(* IEC 61131-3 sources: PLCGen/codesys_service/bank/st_part4, 20 files *)

(* ---- E01_Filling.st ---- *)
(* Q01 Automated Filling Line Control - reference solution for test-case validation *)
FUNCTION_BLOCK E01_Filling
VAR_INPUT
    bottleSensor          : BOOL;
    cleaningConfirmButton : BOOL;
    fillingConfirmButton  : BOOL;
    cappingConfirmButton  : BOOL;
    packingConfirmButton  : BOOL;
    finishedButton        : BOOL;
END_VAR
VAR_OUTPUT
    Pump_Motor       : BOOL;
    Filling_Valve    : BOOL;
    Capping_Machine  : BOOL;
    Packing_Machine  : BOOL;
    Completion_Light : BOOL;
END_VAR
VAR
    step : INT := 0;   (* 0 idle, 1 cleaning, 2 filling, 3 capping, 4 packing, 5 done *)
    prevBottle      : BOOL;
    prevCleaning    : BOOL;
    prevFilling     : BOOL;
    prevCapping     : BOOL;
    prevPacking     : BOOL;
    prevFinished    : BOOL;
END_VAR

(* confirmation is edge-triggered: a button that is already held when its
   step is reached has no rising edge and must not confirm the step *)
IF step = 0 AND bottleSensor AND NOT prevBottle THEN
    step := 1;
ELSIF step = 1 AND cleaningConfirmButton AND NOT prevCleaning THEN
    step := 2;
ELSIF step = 2 AND fillingConfirmButton AND NOT prevFilling THEN
    step := 3;
ELSIF step = 3 AND cappingConfirmButton AND NOT prevCapping THEN
    step := 4;
ELSIF step = 4 AND packingConfirmButton AND NOT prevPacking THEN
    step := 5;
ELSIF step = 5 AND finishedButton AND NOT prevFinished THEN
    step := 0;
END_IF;

Pump_Motor       := step = 1;
Filling_Valve    := step = 2;
Capping_Machine  := step = 3;
Packing_Machine  := step = 4;
Completion_Light := step = 5;

prevBottle   := bottleSensor;
prevCleaning := cleaningConfirmButton;
prevFilling  := fillingConfirmButton;
prevCapping  := cappingConfirmButton;
prevPacking  := packingConfirmButton;
prevFinished := finishedButton;

(* ---- E02_DualEdge.st ---- *)
(* Q02 Dual-Word Edge Detection - reference solution *)
FUNCTION_BLOCK E02_DualEdge
VAR_INPUT
    value : DWORD;
END_VAR
VAR_OUTPUT
    hasChanged      : BOOL;
    hasRisingEdges  : BOOL;
    risingBits      : DWORD;
    noOfRisingBits  : USINT;
    hasFallingEdges : BOOL;
    fallingBits     : DWORD;
    noOfFallingBits : USINT;
END_VAR
VAR
    prev : DWORD;
    i    : INT;
    r    : DWORD;
    f    : DWORD;
END_VAR

risingBits  := value AND NOT prev;
fallingBits := prev AND NOT value;
hasChanged  := value <> prev;
hasRisingEdges  := risingBits <> 0;
hasFallingEdges := fallingBits <> 0;

(* popcount without SHL: shift right by division, which keeps the
   implementation portable and works in the simulator *)
r := risingBits;
f := fallingBits;
noOfRisingBits  := 0;
noOfFallingBits := 0;
FOR i := 0 TO 31 DO
    IF (r MOD 2) <> 0 THEN
        noOfRisingBits := noOfRisingBits + 1;
    END_IF;
    IF (f MOD 2) <> 0 THEN
        noOfFallingBits := noOfFallingBits + 1;
    END_IF;
    r := r / 2;
    f := f / 2;
END_FOR;

prev := value;

(* ---- E03_Hysteresis.st ---- *)
(* Q03 Alarm Handling - reference solution (used only to validate the test cases)
   Note: status codes are written in decimal (32769 = 16#8001, 32770 = 16#8002)
   because the offline simulator (st_sim) does not support typed literals. *)
FUNCTION_BLOCK E03_Hysteresis
VAR_INPUT
    Value      : REAL;
    hiLevel    : REAL;
    loLevel    : REAL;
    hystWindow : REAL;
END_VAR
VAR_OUTPUT
    hiAlarm : BOOL;
    loAlarm : BOOL;
    error   : BOOL;
    status  : WORD;
END_VAR

IF loLevel >= hiLevel THEN
    error  := TRUE;
    status := 32769;
ELSIF hystWindow >= hiLevel - loLevel THEN
    error  := TRUE;
    status := 32770;
ELSE
    error  := FALSE;
    status := 0;
    (* high alarm with hysteresis *)
    IF Value > hiLevel THEN
        hiAlarm := TRUE;
    ELSIF Value < hiLevel - hystWindow THEN
        hiAlarm := FALSE;
    END_IF;
    (* low alarm with hysteresis *)
    IF Value < loLevel THEN
        loAlarm := TRUE;
    ELSIF Value > loLevel + hystWindow THEN
        loAlarm := FALSE;
    END_IF;
END_IF;

(* ---- E04_JamPump.st ---- *)
(* Q04 Jam Pump Debouncing and Runtime Maintenance - reference solution
   Unit convention: TIME inputs in ms, LTIME output in ns (IEC 61131-3). *)
FUNCTION_BLOCK E04_JamPump
VAR_INPUT
    VISCOSITY_OK    : BOOL;
    PASTE_E_STOP_NC : BOOL;
    DebounceTime    : TIME;
    CycleTime       : TIME;
END_VAR
VAR_OUTPUT
    VFD_RUN          : BOOL;
    PUMP_MAINT_DUE   : BOOL;
    PUMP_RUNTIME_ACC : LTIME;
END_VAR
VAR
    debT    : TON;     (* real elapsed time, scan-clock driven *)
    accMs   : ULINT;   (* ms, per the team convention *)
END_VAR

(* VISCOSITY_OK must hold continuously for DebounceTime (real elapsed time) *)
debT(IN := VISCOSITY_OK AND PASTE_E_STOP_NC, PT := DebounceTime);
VFD_RUN := debT.Q AND PASTE_E_STOP_NC;

IF VFD_RUN THEN
    accMs := accMs + UDINT_TO_ULINT(TIME_TO_UDINT(CycleTime));
    PUMP_RUNTIME_ACC := ULINT_TO_LTIME(accMs);
END_IF;

IF accMs >= 1800000000 THEN   (* 500 h in ms *)
    PUMP_MAINT_DUE := TRUE;
END_IF;

(* ---- E05_WeldGap.st ---- *)
(* Q05 Weld Gap Alarm and Startup Inhibition - reference solution *)
FUNCTION_BLOCK E05_WeldGap
VAR_INPUT
    Gap_Exceeded   : BOOL;
    Weld_E_Stop_NC : BOOL;
    DebounceTime   : TIME;
END_VAR
VAR_OUTPUT
    Operator_Alert        : BOOL;
    Weld_Soft_Start_Active: BOOL;
END_VAR
VAR
    initTimer : TON;
    debTimer  : TON;
    initDone  : BOOL;
END_VAR

initTimer(IN := Weld_E_Stop_NC AND NOT initDone, PT := T#5S);
IF initTimer.Q THEN
    initDone := TRUE;
END_IF;

IF NOT Weld_E_Stop_NC THEN
    Operator_Alert := FALSE;
    Weld_Soft_Start_Active := FALSE;
    debTimer(IN := FALSE, PT := DebounceTime);
ELSIF NOT initDone THEN
    Operator_Alert := FALSE;
    Weld_Soft_Start_Active := TRUE;
    debTimer(IN := FALSE, PT := DebounceTime);
ELSE
    Weld_Soft_Start_Active := FALSE;
    debTimer(IN := Gap_Exceeded, PT := DebounceTime);
    Operator_Alert := debTimer.Q;
END_IF;

(* ---- E06_Blower.st ---- *)
(* Q06 Aeration Blower Delayed Start - reference solution *)
FUNCTION_BLOCK E06_Blower
VAR_INPUT
    DO_LOW               : BOOL;
    AERATION_E_STOP_NC   : BOOL;
END_VAR
VAR_OUTPUT
    BLOWER_RUN                  : BOOL;
    AERATION_BLOWER_CYCLE_COUNT : UINT;
END_VAR
VAR
    startTimer : TON;
    prevRun    : BOOL;
END_VAR

startTimer(IN := DO_LOW AND AERATION_E_STOP_NC, PT := T#5S);
BLOWER_RUN := startTimer.Q;

IF BLOWER_RUN AND NOT prevRun THEN
    AERATION_BLOWER_CYCLE_COUNT := AERATION_BLOWER_CYCLE_COUNT + 1;
END_IF;
prevRun := BLOWER_RUN;

(* ---- H01_Proportion.st ---- *)
(* Q15 Material Proportioning Process Control - reference solution for test-case validation *)
FUNCTION_BLOCK H01_Proportion
VAR_INPUT
    estop           : BOOL;
    opeMode         : BOOL;
    valveAStart     : BOOL;
    valveBStart     : BOOL;
    valveCStart     : BOOL;
    valveDStart     : BOOL;
    mixMotorStart   : BOOL;
    autoStart       : BOOL;
    processMode     : BOOL;
    levelSensor     : INT;
    mixMotorComplete: BOOL;
END_VAR
VAR_OUTPUT
    valveARun   : BOOL;
    valveBRun   : BOOL;
    valveCRun   : BOOL;
    valveDRun   : BOOL;
    mixMotorRun : BOOL;
END_VAR
VAR
    step : INT := 0;
    pA : BOOL;
    pB : BOOL;
    pC : BOOL;
    pD : BOOL;
    pM : BOOL;
END_VAR

IF NOT estop THEN
    valveARun := FALSE;
    valveBRun := FALSE;
    valveCRun := FALSE;
    valveDRun := FALSE;
    mixMotorRun := FALSE;
    step := 0;
ELSIF NOT opeMode THEN
    step := 0;
    IF valveAStart AND NOT pA THEN valveARun := NOT valveARun; END_IF;
    IF valveBStart AND NOT pB THEN valveBRun := NOT valveBRun; END_IF;
    IF valveCStart AND NOT pC THEN valveCRun := NOT valveCRun; END_IF;
    IF valveDStart AND NOT pD THEN valveDRun := NOT valveDRun; END_IF;
    IF mixMotorStart AND NOT pM THEN mixMotorRun := NOT mixMotorRun; END_IF;
ELSE
    IF step = 0 THEN
        valveARun := FALSE;
    valveBRun := FALSE;
    valveCRun := FALSE;
    valveDRun := FALSE;
    mixMotorRun := FALSE;
        IF autoStart THEN step := 1; END_IF;
    END_IF;
    IF step = 1 THEN
        valveARun := TRUE;
        IF levelSensor >= 50 THEN valveARun := FALSE; step := 2; END_IF;
    END_IF;
    IF step = 2 THEN
        valveBRun := TRUE;
        IF levelSensor >= 80 THEN
            valveBRun := FALSE;
            IF processMode THEN step := 3; ELSE step := 4; END_IF;
        END_IF;
    END_IF;
    IF step = 3 THEN
        valveCRun := TRUE;
        IF levelSensor >= 100 THEN valveCRun := FALSE; step := 4; END_IF;
    END_IF;
    IF step = 4 THEN
        mixMotorRun := TRUE;
        IF mixMotorComplete THEN mixMotorRun := FALSE; valveDRun := TRUE; step := 5; END_IF;
    END_IF;
END_IF;
pA := valveAStart;
pB := valveBStart;
pC := valveCStart;
pD := valveDStart;
pM := mixMotorStart;

(* ---- H02_FlexProcess.st ---- *)
(* Q16 Flexible Processing Control - reference solution *)
FUNCTION_BLOCK H02_FlexProcess
VAR_INPUT
    processLength   : USINT;
    sensor1         : BOOL;
    sensor2         : BOOL;
    sensor3         : BOOL;
    sensor4         : BOOL;
    sensor5         : BOOL;
    station1Start   : BOOL;
    station2Complete: BOOL;
    station3Complete: BOOL;
    station4Complete: BOOL;
    processSequence : ARRAY[1..8] OF USINT;
END_VAR
VAR_OUTPUT
    conveyorLeft  : BOOL;
    conveyorRight : BOOL;
END_VAR
VAR
    idx     : USINT;      (* active entry, 0 = not started *)
    cur     : USINT;      (* station the product is at, 0 = in transit *)
    target  : USINT;
    moving  : BOOL;
    atTarget: BOOL;
    done    : BOOL;
END_VAR

conveyorLeft := FALSE;
conveyorRight := FALSE;

(* Station tracking.  The carriage position is latched when it arrives: the
   sensors alone cannot be used, because the sensor of the station just left
   drops while the carriage is in transit, which would erase the direction
   needed for the next leg. *)
IF sensor1 THEN cur := 1; END_IF;
IF sensor2 THEN cur := 2; END_IF;
IF sensor3 THEN cur := 3; END_IF;
IF sensor4 THEN cur := 4; END_IF;
IF sensor5 THEN cur := 5; END_IF;

IF idx = 0 AND sensor1 AND station1Start THEN
    idx := 1;
    moving := TRUE;
    cur := 1;                                (* latched, not re-read from sensor1 *)
END_IF;

IF idx > 0 THEN
    target := processSequence[idx];
    atTarget := (cur = target);

    IF moving AND atTarget THEN
        moving := FALSE;                     (* arrived: stop *)
        conveyorLeft := FALSE;
        conveyorRight := FALSE;
        cur := target;                       (* latch: the sensor may drop *)
    END_IF;

    IF NOT moving AND atTarget THEN
        done := FALSE;
        IF target = 2 THEN
            done := station2Complete;
        ELSIF target = 3 THEN
            done := station3Complete;
        ELSIF target = 4 THEN
            done := station4Complete;
        END_IF;
        IF done AND idx < processLength THEN
            idx := idx + 1;
            moving := TRUE;
        END_IF;
    END_IF;

    IF moving THEN
        target := processSequence[idx];
        IF target > cur THEN
            conveyorRight := TRUE;
        ELSIF target < cur THEN
            conveyorLeft := TRUE;
        END_IF;
    END_IF;
END_IF;

(* ---- H03_RecipeMgr.st ---- *)
TYPE ST_Recipe :
STRUCT
    recipeID              : INT;
    ingredientType        : INT;
    ingredientRatio       : REAL;
    productionTemperature : REAL;
END_STRUCT
END_TYPE

(* Q17 Recipe Management System - reference solution *)
FUNCTION_BLOCK H03_RecipeMgr
VAR_INPUT
    addRecipe    : BOOL;
    deleteRecipe : BOOL;
    modifyRecipe : BOOL;
    queryRecipe  : BOOL;
    recipeIn     : ST_Recipe;
END_VAR
VAR_OUTPUT
    recipeAdded       : BOOL;
    recipeDeleted     : BOOL;
    recipeModified    : BOOL;
    recipeQueryResult : ST_Recipe;
    error             : BOOL;
    status            : WORD;
END_VAR
VAR_IN_OUT
    recipe : ARRAY[1..10] OF ST_Recipe;
END_VAR
VAR
    i    : INT;
    slot : INT;
    free : INT;
END_VAR

recipeAdded := FALSE;
recipeDeleted := FALSE;
recipeModified := FALSE;
error := FALSE;
status := 16#0000;

slot := 0;
free := 0;
FOR i := 10 TO 1 BY -1 DO
    IF recipe[i].recipeID = recipeIn.recipeID THEN
        slot := i;
    END_IF;
    IF recipe[i].recipeID = 0 THEN
        free := i;
    END_IF;
END_FOR;

IF queryRecipe THEN
    IF slot = 0 THEN
        error := TRUE;
        status := 16#8001;
    ELSE
        recipeQueryResult := recipe[slot];
    END_IF;
ELSIF addRecipe THEN
    IF slot <> 0 THEN
        error := TRUE;
        status := 16#8002;
    ELSIF free = 0 THEN
        error := TRUE;
        status := 16#8003;
    ELSE
        recipe[free] := recipeIn;
        recipeAdded := TRUE;
    END_IF;
ELSIF deleteRecipe THEN
    IF slot = 0 THEN
        error := TRUE;
        status := 16#8004;
    ELSE
        recipe[slot].recipeID := 0;
        recipeDeleted := TRUE;
    END_IF;
ELSIF modifyRecipe THEN
    IF slot = 0 THEN
        error := TRUE;
        status := 16#8005;
    ELSE
        recipe[slot] := recipeIn;
        recipeModified := TRUE;
    END_IF;
END_IF;

(* ---- H04_FIFO.st ---- *)
(* H04 FIFO Queue - reference solution.
   The interface uses VARIANT in the task; this reference uses a concrete
   array so that it can be compiled and tested in the harness.
   Buffer capacity is 8 (ARRAY[0..7] OF DINT), the convention settled with
   Part 2; the test cases assume exactly this. *)
FUNCTION_BLOCK H04_FIFO
VAR_INPUT
    enqueue : BOOL;
    dequeue : BOOL;
    reset   : BOOL;
END_VAR
VAR_OUTPUT
    elementCount : DINT;
    status       : WORD;
END_VAR
VAR_IN_OUT
    item   : DINT;
    buffer : ARRAY[0..7] OF DINT;
END_VAR
VAR
    head : DINT := 0;
    tail : DINT := 0;
    cap  : DINT := 8;   (* ARRAY[0..7] *)
    prevEnq : BOOL;
    prevDeq : BOOL;
    enqEdge : BOOL;
    deqEdge : BOOL;
END_VAR

status := 16#0000;
enqEdge := enqueue AND NOT prevEnq;
deqEdge := dequeue AND NOT prevDeq;
prevEnq := enqueue;
prevDeq := dequeue;

IF reset THEN
    head := 0;
    tail := 0;
    elementCount := 0;
ELSIF enqEdge THEN
    IF elementCount >= cap THEN
        status := 16#8002;
    ELSE
        buffer[tail] := item;
        tail := tail + 1;
        IF tail >= cap THEN
            tail := 0;
        END_IF;
        elementCount := elementCount + 1;
    END_IF;
ELSIF deqEdge THEN
    IF elementCount <= 0 THEN
        status := 16#8001;
    ELSE
        item := buffer[head];
        head := head + 1;
        IF head >= cap THEN
            head := 0;
        END_IF;
        elementCount := elementCount - 1;
    END_IF;
END_IF;

(* ---- H05_MechArm.st ---- *)
(* Q19 Mechanical Arm Control - reference solution for test-case validation *)
FUNCTION_BLOCK H05_MechArm
VAR_INPUT
    ManualMode        : BOOL;
    SingleStepMode    : BOOL;
    SingleCycleMode   : BOOL;
    ContinuousMode    : BOOL;
    EmergencyStop     : BOOL;
    Start             : BOOL;
    DownButton        : BOOL;
    UpButton          : BOOL;
    LeftButton        : BOOL;
    RightButton       : BOOL;
    GripButton        : BOOL;
    ReleaseButton     : BOOL;
    DownLimitSwitch   : BOOL;
    UpLimitSwitch     : BOOL;
    LeftLimitSwitch   : BOOL;
    RightLimitSwitch  : BOOL;
    GripLimitSwitch   : BOOL;
    ReleaseLimitSwitch: BOOL;
END_VAR
VAR_OUTPUT
    MoveDown        : BOOL;
    MoveUp          : BOOL;
    MoveLeft        : BOOL;
    MoveRight       : BOOL;
    ActivateGrip    : BOOL;
    ActivateRelease : BOOL;
END_VAR
VAR
    step    : INT := 0;   (* 0 idle at top-left; 1 down 2 grip 3 up 4 right 5 down 6 release 7 up 8 left *)
    active  : BOOL;       (* current step is being executed *)
    pStart  : BOOL;
    startEdge : BOOL;
    stepDone : BOOL;
END_VAR

startEdge := Start AND NOT pStart;
pStart := Start;

MoveDown := FALSE;
MoveUp := FALSE;
MoveLeft := FALSE;
MoveRight := FALSE;
ActivateGrip := FALSE;
ActivateRelease := FALSE;

IF NOT EmergencyStop THEN
    active := FALSE;
    step := 0;
ELSIF ManualMode THEN
    active := FALSE;
    step := 0;
    MoveDown := DownButton AND NOT DownLimitSwitch;
    MoveUp := UpButton AND NOT UpLimitSwitch;
    MoveLeft := LeftButton AND NOT LeftLimitSwitch;
    MoveRight := RightButton AND NOT RightLimitSwitch;
    ActivateGrip := GripButton AND NOT GripLimitSwitch;
    ActivateRelease := ReleaseButton AND NOT ReleaseLimitSwitch;
ELSE
    (* start a step when idle *)
    IF NOT active THEN
        IF startEdge THEN
            IF step = 0 OR step = 8 THEN
                step := 1;
            ELSE
                step := step + 1;
            END_IF;
            active := TRUE;
        END_IF;
    END_IF;

    IF active THEN
        stepDone := FALSE;
        IF step = 1 OR step = 5 THEN
            MoveDown := NOT DownLimitSwitch;
            stepDone := DownLimitSwitch;
        ELSIF step = 2 THEN
            ActivateGrip := NOT GripLimitSwitch;
            stepDone := GripLimitSwitch;
        ELSIF step = 3 OR step = 7 THEN
            MoveUp := NOT UpLimitSwitch;
            stepDone := UpLimitSwitch;
        ELSIF step = 4 THEN
            MoveRight := NOT RightLimitSwitch;
            stepDone := RightLimitSwitch;
        ELSIF step = 6 THEN
            ActivateRelease := NOT ReleaseLimitSwitch;
            stepDone := ReleaseLimitSwitch;
        ELSIF step = 8 THEN
            MoveLeft := NOT LeftLimitSwitch;
            stepDone := LeftLimitSwitch;
        END_IF;

        IF stepDone THEN
            IF SingleStepMode THEN
                active := FALSE;                 (* wait for next Start *)
            ELSIF step < 8 THEN
                step := step + 1;                (* cycle modes: chain to next step *)
            ELSE
                step := 0;
                IF NOT ContinuousMode THEN
                    active := FALSE;             (* single cycle: stop at home *)
                ELSE
                    step := 1;                   (* continuous: restart *)
                END_IF;
            END_IF;
        END_IF;
    END_IF;
END_IF;

(* ---- H06_Production.st ---- *)
(* Q20 Production Control - reference solution for test-case validation *)
FUNCTION_BLOCK H06_Production
VAR_INPUT
    Mode           : BOOL;
    ForwardButton  : BOOL;
    ReverseButton  : BOOL;
    SensorFeed     : BOOL;
    SensorWash     : BOOL;
    SensorWeight   : BOOL;
    SensorFiring   : BOOL;
    SensorOutput   : BOOL;
    washComplete   : BOOL;
    weightComplete : BOOL;
    weight         : REAL;
    firingComplete : BOOL;
END_VAR
VAR_OUTPUT
    MotorForward    : BOOL;
    MotorReverse    : BOOL;
    kick            : BOOL;
    CompletionLight : BOOL;
    firingTemp      : REAL;
END_VAR
VAR
    step : INT := 0;
    (* 0 idle, 1 feed->wash, 2 at wash, 3 wash->weight, 4 at weight, 5 rejected,
       6 weight->firing, 7 at firing, 8 firing->output, 9 at output *)
END_VAR

IF NOT Mode THEN
    MotorForward := ForwardButton AND NOT ReverseButton;
    MotorReverse := ReverseButton AND NOT ForwardButton;
    kick := FALSE;
    CompletionLight := FALSE;
    step := 0;
ELSE
    MotorReverse := FALSE;
    kick := FALSE;
    IF step = 0 AND SensorFeed THEN
        step := 1;
    ELSIF step = 1 AND SensorWash THEN
        step := 2;
    ELSIF step = 2 AND washComplete THEN
        step := 3;
    ELSIF step = 3 AND SensorWeight THEN
        step := 4;
    ELSIF step = 4 AND weightComplete THEN
        IF weight >= 100.0 AND weight <= 200.0 THEN
            firingTemp := 500.0 + (weight - 100.0) * 0.5;
            step := 6;
        ELSE
            kick := TRUE;
            step := 5;
        END_IF;
    ELSIF step = 5 AND NOT SensorWeight THEN
        step := 0;
    ELSIF step = 6 AND SensorFiring THEN
        step := 7;
    ELSIF step = 7 AND firingComplete THEN
        step := 8;
    ELSIF step = 8 AND SensorOutput THEN
        step := 9;
    ELSIF step = 9 AND NOT SensorOutput THEN
        step := 0;
    END_IF;
    MotorForward := step = 1 OR step = 3 OR step = 6 OR step = 8;
    CompletionLight := step = 9;
END_IF;

(* ---- M01_PumpSwitch.st ---- *)
TYPE ST_Pump :
STRUCT
    priority  : INT;
    selection : BOOL;
    RunComd   : BOOL;
END_STRUCT
END_TYPE

(* Q07 Multi-Pump Switching Control System - reference solution *)
FUNCTION_BLOCK M01_PumpSwitch
VAR_INPUT
    mode  : BOOL;
    start : BOOL;
    stop  : BOOL;
END_VAR
VAR_IN_OUT
    pumpGroup : ARRAY[1..5] OF ST_Pump;
END_VAR
VAR
    i, j, best, bestIdx, picked : INT;
    chosen : ARRAY[1..5] OF BOOL;
    running : BOOL;
END_VAR

IF stop THEN
    FOR i := 1 TO 5 DO
        pumpGroup[i].RunComd := FALSE;
    END_FOR;
    running := FALSE;
ELSIF start THEN
    running := TRUE;
END_IF;

IF running THEN
    IF NOT mode THEN
        (* manual: run exactly the selected pumps *)
        FOR i := 1 TO 5 DO
            pumpGroup[i].RunComd := pumpGroup[i].selection;
        END_FOR;
    ELSE
        (* automatic: three highest priorities run, two stand by *)
        FOR i := 1 TO 5 DO
            chosen[i] := FALSE;
        END_FOR;
        FOR picked := 1 TO 3 DO
            bestIdx := 0;
            FOR j := 1 TO 5 DO
                IF NOT chosen[j] THEN
                    IF bestIdx = 0 THEN
                        bestIdx := j;
                        best := pumpGroup[j].priority;
                    ELSIF pumpGroup[j].priority > best THEN
                        bestIdx := j;
                        best := pumpGroup[j].priority;
                    END_IF;
                END_IF;
            END_FOR;
            IF bestIdx > 0 THEN
                chosen[bestIdx] := TRUE;
            END_IF;
        END_FOR;
        FOR i := 1 TO 5 DO
            pumpGroup[i].RunComd := chosen[i];
        END_FOR;
    END_IF;
END_IF;

(* ---- M02_AnalogBatch.st ---- *)
TYPE ST_AnalogChannel :
STRUCT
    enable        : BOOL;
    hiLIM         : REAL;
    loLIM         : REAL;
    bipolar       : BOOL;
    measuringMode : INT;
    retVal        : WORD;
    outputValue   : REAL;
END_STRUCT
END_TYPE

(* Q08 Analog Batch Processing - reference solution.
   The task declares ARRAY[*]; this reference fixes the length at 2 so that it
   can be compiled and exercised by the test harness. *)
FUNCTION_BLOCK M02_AnalogBatch
VAR_INPUT
    count : DINT;
END_VAR
VAR_IN_OUT
    analogValues : ARRAY[1..2] OF INT;
    channels     : ARRAY[1..2] OF ST_AnalogChannel;
END_VAR
VAR
    i   : DINT;
    raw : REAL;
END_VAR

FOR i := 1 TO 2 DO
    IF i <= count AND channels[i].enable THEN
        IF channels[i].measuringMode < 0 OR channels[i].measuringMode > 2 THEN
            channels[i].retVal := 16#8001;
        ELSIF channels[i].hiLIM <= channels[i].loLIM THEN
            channels[i].retVal := 16#8002;
        ELSE
            channels[i].retVal := 16#0000;
            raw := INT_TO_REAL(analogValues[i]);
            IF channels[i].measuringMode = 0 THEN
                IF channels[i].bipolar THEN
                    channels[i].outputValue := channels[i].loLIM
                        + (raw + 27648.0) / 55296.0 * (channels[i].hiLIM - channels[i].loLIM);
                ELSE
                    channels[i].outputValue := channels[i].loLIM
                        + raw / 27648.0 * (channels[i].hiLIM - channels[i].loLIM);
                END_IF;
            ELSIF channels[i].measuringMode = 1 THEN
                channels[i].outputValue := raw / 10.0;
            ELSE
                channels[i].outputValue := raw / 100.0;
            END_IF;
        END_IF;
    END_IF;
END_FOR;

(* ---- M03_MovingAvg.st ---- *)
(* Q09 Calculate Moving Average - reference solution *)
FUNCTION_BLOCK M03_MovingAvg
VAR_INPUT
    cyclicExecution : BOOL;
    trigger         : BOOL;
    value           : LREAL;
    windowSize      : INT;
    reset           : BOOL;
END_VAR
VAR_OUTPUT
    average            : LREAL;
    windowSizeReached  : BOOL;
    error              : BOOL;
    status             : WORD;
END_VAR
VAR
    buf   : ARRAY[0..99] OF LREAL;
    count : INT;
    head  : INT;
    sum   : LREAL;
    prevTrig : BOOL;
    doRead : BOOL;
    i : INT;
END_VAR

(* Validation first: an out-of-range window must not touch the buffer. *)
IF windowSize < 1 OR windowSize > 100 THEN
    error := TRUE;
    status := 16#8200;
    average := 0;
    windowSizeReached := FALSE;
    prevTrig := trigger;
ELSIF reset THEN
    (* reset clears the window and the result *)
    count := 0;
    head := 0;
    sum := 0;
    average := 0;
    windowSizeReached := FALSE;
    error := FALSE;
    status := 16#0000;
    prevTrig := trigger;
ELSE
    error := FALSE;
    status := 16#0000;

    IF cyclicExecution THEN
        doRead := TRUE;
    ELSE
        doRead := trigger AND NOT prevTrig;
    END_IF;
    prevTrig := trigger;

    IF doRead THEN
        IF count < windowSize THEN
            buf[head] := value;
            sum := sum + value;
            count := count + 1;
        ELSE
            sum := sum - buf[head];
            buf[head] := value;
            sum := sum + value;
        END_IF;
        head := head + 1;
        IF head >= windowSize THEN
            head := 0;
        END_IF;
    END_IF;

    IF count > 0 THEN
        average := sum / INT_TO_LREAL(count);
    ELSE
        average := 0;
    END_IF;
    windowSizeReached := count >= windowSize;
END_IF;

(* ---- M04_TempCtrl.st ---- *)
(* Q10 Temperature Logic Control - reference solution *)
FUNCTION_BLOCK M04_TempCtrl
VAR_INPUT
    TemperatureSensorInput : REAL;
    SetTemperature         : REAL;
END_VAR
VAR_OUTPUT
    CurrentTemperature : REAL;
    SetTempDisplay     : REAL;
    HeaterStatus       : BOOL;
    OverheatProtection : BOOL;
    HeaterOutput       : BOOL;
END_VAR
VAR
    runTimer  : TON;
    coolTimer : TON;
    sensorFault : BOOL;
END_VAR

CurrentTemperature := TemperatureSensorInput;
SetTempDisplay := SetTemperature;
sensorFault := TemperatureSensorInput < 0.0 OR TemperatureSensorInput > 100.0;

runTimer(IN := HeaterOutput, PT := T#5S);
IF runTimer.Q THEN
    OverheatProtection := TRUE;
END_IF;

coolTimer(IN := OverheatProtection, PT := T#3S);
IF coolTimer.Q THEN
    OverheatProtection := FALSE;
END_IF;

IF sensorFault OR OverheatProtection THEN
    HeaterOutput := FALSE;
ELSIF TemperatureSensorInput < SetTemperature THEN
    HeaterOutput := TRUE;
ELSE
    HeaterOutput := FALSE;
END_IF;

HeaterStatus := HeaterOutput;

(* ---- M05_ProdLine.st ---- *)
(* Q11 Automated Production Line Control - reference solution for test-case validation *)
FUNCTION_BLOCK M05_ProdLine
VAR_INPUT
    Mode          : BOOL;
    ForwardButton : BOOL;
    ReverseButton : BOOL;
    SensorA       : BOOL;
    SensorB       : BOOL;
    SensorC       : BOOL;
    ButtonA       : BOOL;
    ButtonB       : BOOL;
    ButtonC       : BOOL;
END_VAR
VAR_OUTPUT
    MotorForward    : BOOL;
    MotorReverse    : BOOL;
    CompletionLight : BOOL;
END_VAR
VAR
    step : INT := 0;  (* 0 wait at A, 1 move A->B, 2 wait at B, 3 move B->C, 4 at C, 5 done *)
    prevA : BOOL;
    prevB : BOOL;
    prevC : BOOL;
    shownStep : INT := 0;   (* the step whose outputs are being driven *)
END_VAR

IF NOT Mode THEN
    (* manual: interlocked jog *)
    MotorForward := ForwardButton AND NOT ReverseButton;
    MotorReverse := ReverseButton AND NOT ForwardButton;
    CompletionLight := FALSE;
    step := 0;
ELSE
    (* Automatic mode.  The motor outputs are assigned inside each step branch and
       cleared in the same scan a transition happens, so the output of a newly
       entered step only appears from the next scan onwards.
       Station buttons are edge-triggered: a button already held when the carriage
       arrives has no rising edge and must not release it. *)
    MotorReverse := FALSE;

    IF step = 0 THEN
        MotorForward := FALSE;
        IF SensorA AND ButtonA AND NOT prevA THEN
            step := 1;
        END_IF;
    ELSIF step = 1 THEN
        MotorForward := TRUE;
        IF SensorB THEN
            MotorForward := FALSE;
            step := 2;
        END_IF;
    ELSIF step = 2 THEN
        MotorForward := FALSE;
        IF ButtonB AND NOT prevB THEN
            step := 3;
        END_IF;
    ELSIF step = 3 THEN
        MotorForward := TRUE;
        IF SensorC THEN
            MotorForward := FALSE;
            step := 4;
        END_IF;
    ELSE
        MotorForward := FALSE;
        IF ButtonC AND NOT prevC THEN
            CompletionLight := TRUE;
        END_IF;
        IF NOT SensorC THEN
            CompletionLight := FALSE;
            step := 0;
        END_IF;
    END_IF;

    prevA := ButtonA;
    prevB := ButtonB;
    prevC := ButtonC;
END_IF;

(* ---- M06_SlabThick.st ---- *)
(* Q12 Slab Thickness Alarm and Fault History - reference solution
   Unit convention: CycleTime in ms, Slab_Runtime_Accumulator in ms (LTIME). *)
FUNCTION_BLOCK M06_SlabThick
VAR_INPUT
    THICKNESS_FAULT        : BOOL;
    THICKNESS_SIGNAL_VALID : BOOL;
    CUTTING_RUN            : BOOL;
    FaultTimestamp         : DINT;
    CycleTime              : TIME;
END_VAR
VAR_OUTPUT
    THICKNESS_ALARM          : BOOL;
    Slab_Fault_Counter       : UINT;
    Slab_Runtime_Accumulator : LTIME;
    Slab_Fault_History       : ARRAY[0..4] OF DINT;
END_VAR
VAR
    holdT    : TON;     (* real elapsed time, scan-clock driven *)
    accMs    : ULINT;   (* ms, per the team convention *)
    prevFlt  : BOOL;
    i        : INT;
END_VAR

IF NOT THICKNESS_SIGNAL_VALID THEN
    THICKNESS_ALARM := FALSE;
    holdT(IN := FALSE, PT := T#500MS);
    prevFlt := FALSE;
ELSE
    IF THICKNESS_FAULT AND NOT prevFlt THEN
        (* new fault: count and record *)
        Slab_Fault_Counter := Slab_Fault_Counter + 1;
        FOR i := 4 TO 1 BY -1 DO
            Slab_Fault_History[i] := Slab_Fault_History[i-1];
        END_FOR;
        Slab_Fault_History[0] := FaultTimestamp;
        THICKNESS_ALARM := TRUE;
        holdT(IN := TRUE, PT := T#500MS);
    END_IF;
    prevFlt := THICKNESS_FAULT;

    IF THICKNESS_ALARM THEN
        (* restart the 500 ms window whenever the fault is still present *)
        holdT(IN := NOT THICKNESS_FAULT, PT := T#500MS);
        IF holdT.Q THEN
            THICKNESS_ALARM := FALSE;
        END_IF;
    END_IF;

    IF CUTTING_RUN AND NOT THICKNESS_FAULT THEN
        accMs := accMs + UDINT_TO_ULINT(TIME_TO_UDINT(CycleTime));
        Slab_Runtime_Accumulator := ULINT_TO_LTIME(accMs);
    END_IF;
END_IF;

(* ---- M07_HVAC.st ---- *)
(* Q13 Office HVAC Multi-mode Energy-Saving Control - reference solution *)
FUNCTION_BLOCK M07_HVAC
VAR_INPUT
    OCCUPANCY_DETECTED : BOOL;
    ENERGY_SAVING_MODE : BOOL;
    HVAC_MODE_SELECTOR : INT;
END_VAR
VAR_OUTPUT
    SUPPLY_FAN_RUN       : BOOL;
    TEMP_SETPOINT_ADJUST : INT;
END_VAR
VAR
    startTimer : TON;
END_VAR

startTimer(IN := OCCUPANCY_DETECTED AND HVAC_MODE_SELECTOR <> 3, PT := T#30S);
SUPPLY_FAN_RUN := startTimer.Q;

IF HVAC_MODE_SELECTOR = 3 THEN
    TEMP_SETPOINT_ADJUST := 4;
ELSIF OCCUPANCY_DETECTED THEN
    TEMP_SETPOINT_ADJUST := 0;
ELSIF HVAC_MODE_SELECTOR = 1 THEN
    TEMP_SETPOINT_ADJUST := 1;
ELSIF HVAC_MODE_SELECTOR = 2 THEN
    TEMP_SETPOINT_ADJUST := 4;
ELSIF ENERGY_SAVING_MODE THEN
    TEMP_SETPOINT_ADJUST := 3;
ELSE
    TEMP_SETPOINT_ADJUST := 2;
END_IF;

(* ---- M08_IPv4.st ---- *)
(* Q14 IPv4 Parsing with Format and Range Checks - reference solution *)
FUNCTION_BLOCK M08_IPv4
VAR_INPUT
    ipText : STRING(254);
END_VAR
VAR_OUTPUT
    ipValue : UDINT;
END_VAR
VAR
    i, n, segCount, digits, segVal : INT;
    ch : BYTE;
    acc : UDINT;
    ok : BOOL;
END_VAR

ipValue := 0;
acc := 0;
segCount := 0;
digits := 0;
segVal := 0;
ok := TRUE;
(* LEN avoids both WHILE and ADR: the simulator supports the Standard string
   functions and direct 1-based indexing of a STRING *)
n := LEN(ipText);

IF n > 0 THEN
FOR i := 1 TO n DO
    ch := ipText[i];
    IF ch >= 48 AND ch <= 57 THEN
        segVal := segVal * 10 + (BYTE_TO_INT(ch) - 48);
        digits := digits + 1;
        IF digits > 3 OR segVal > 255 THEN
            ok := FALSE;
        END_IF;
    ELSIF ch = 46 THEN
        IF digits = 0 THEN
            ok := FALSE;
        END_IF;
        acc := acc * 256 + INT_TO_UDINT(segVal);
        segCount := segCount + 1;
        segVal := 0;
        digits := 0;
        IF segCount > 3 THEN
            ok := FALSE;
        END_IF;
    ELSE
        ok := FALSE;
    END_IF;
END_FOR;
END_IF;

IF digits = 0 THEN
    ok := FALSE;
END_IF;
acc := acc * 256 + INT_TO_UDINT(segVal);
segCount := segCount + 1;

IF ok AND segCount = 4 THEN
    ipValue := acc;
END_IF;
